(* IEC 61131-3 sources: NachHouse_TST/ROOM_API_PILOT/CODEX_BACKUP_BEFORE_SORT_FIX_20260827_0827, 1 file *)

(* ---- 08_COMMAND_ENGINE.ST ---- *)
(* Spracovanie príkazov ADD / DELETE / COPY / SET pre miestnosti. ENG *)

(* Spracuje najviac jeden príkaz, iba ak klient nastavil ApiCommandExecute. *)
FUNCTION ApiProcessRoomCommand : BOOL
VAR
    i             : USINT;     (* Index pri prechode poľom miestností. *)
    configSlot    : USINT;     (* Nájdená alebo voľná pozícia cieľovej konfigurácie. ENG *)
    stateSlot     : USINT;     (* Nájdená alebo voľná pozícia cieľového stavu. ENG *)
    sourceCfgSlot : USINT;     (* Pozícia zdrojovej konfigurácie pri kopírovaní. ENG *)
    sourceStSlot  : USINT;     (* Pozícia zdrojového stavu pri kopírovaní. ENG *)
    maxSort       : UINT;      (* Najvyššie použité predvolené poradie pri pridávaní. ENG *)
    sourceSort    : UINT;      (* Predvolené poradie zdroja pri vkladaní jeho kópie. ENG *)
    resultCode    : USINT;     (* Pracovný návratový kód API_RESULT_*. ENG *)
    resultMessage : STRING[80]; (* Pracovný slovenský text výsledku. *)
    executeChange : BOOL;      (* TRUE iba vtedy, keď sa snapshot skutočne zmenil. ENG *)
END_VAR

(* Bez spúšťacieho príznaku funkcia okamžite skončí bez vedľajších účinkov. *)
ApiProcessRoomCommand := FALSE;
IF NOT ApiCommandExecute THEN
    RETURN;
END_IF;

(* Začiatok dvojfázového handshake: príkaz je prevzatý na spracovanie. ENG *)
ApiProcessRoomCommand := TRUE;
ApiCommandBusy := TRUE;
ApiCommandFinished := FALSE;

(* Presné zopakovanie posledného ClientId + RequestId je idempotentné. ENG *)
IF (ApiCommandRoom.ClientId = ApiLastCommandClientId) AND
   (ApiCommandRoom.RequestId = ApiLastCommandRequestId) AND
   (ApiCommandRoom.RequestId <> 0) THEN

    ApiCommandResult := ApiLastStoredResult;
    ApiInfo.LastCommandResult := ApiLastStoredResult;

ELSE
    (* Predvolené hodnoty pre nový, ešte nespracovaný príkaz. *)
    resultCode := API_RESULT_OK;
    resultMessage := 'OK';
    executeChange := FALSE;

    (* Spoločná kontrola povinných identifikátorov transportu. *)
    IF (ApiCommandRoom.ClientId = '') OR (ApiCommandRoom.RequestId = 0) THEN
        resultCode := API_RESULT_INVALID_ARGUMENT;
        resultMessage := 'Neplatny ClientId alebo RequestId';
    ELSE
        (* Rozdelenie spracovania podľa verejného číselného kódu Action. ENG *)
        CASE ApiCommandRoom.Action OF

            API_ACTION_ADD_ROOM:
                (* ADD: overí cieľ, nájde voľné sloty a vytvorí konfiguráciu aj stav. ENG *)
                IF (ApiCommandRoom.RoomId = 0) OR (ApiCommandRoom.Name = '') THEN
                    resultCode := API_RESULT_INVALID_ARGUMENT;
                    resultMessage := 'Neplatne ID alebo nazov';
                ELSIF ApiFindConfigSlot(ApiCommandRoom.RoomId) <> 0 THEN
                    resultCode := API_RESULT_ALREADY_EXISTS;
                    resultMessage := 'RoomId uz existuje';
                ELSE
                    configSlot := ApiFindFreeConfigSlot();
                    stateSlot := ApiFindFreeStateSlot();
                    IF (configSlot = 0) OR (stateSlot = 0) THEN
                        resultCode := API_RESULT_NO_FREE_SLOT;
                        resultMessage := 'Nie je volny slot';
                    ELSE
                        (* Nová miestnosť sa zaradí za najvyššie existujúce SortDefault. ENG *)
                        maxSort := 0;
                        FOR i := 1 TO C_MAX_ROOMS DO
                            IF ApiConfig.Rooms[i].Used AND
                               (ApiConfig.Rooms[i].SortDefault > maxSort) THEN
                                maxSort := ApiConfig.Rooms[i].SortDefault;
                            END_IF;
                        END_FOR;

                        (* Vytvorenie cieľovej konfigurácie z údajov klienta a predvolenej ikony. *)
                        ApiClearRoomConfig(ApiConfig.Rooms[configSlot]);
                        ApiConfig.Rooms[configSlot].Used := TRUE;
                        ApiConfig.Rooms[configSlot].RoomId := ApiCommandRoom.RoomId;
                        ApiConfig.Rooms[configSlot].Name := ApiCommandRoom.Name;
                        ApiConfig.Rooms[configSlot].ProjectName := ApiCommandRoom.ProjectName;
                        ApiConfig.Rooms[configSlot].IconId := API_DEFAULT_ICON_ID;
                        ApiConfig.Rooms[configSlot].SortDefault := maxSort + 1;

                        (* Vytvorenie samostatného stavového záznamu s testovacími hodnotami. *)
                        ApiClearRoomState(ApiState.Rooms[stateSlot]);
                        ApiState.Rooms[stateSlot].RoomId := ApiCommandRoom.RoomId;
                        ApiState.Rooms[stateSlot].Temperature := API_DEFAULT_TEMPERATURE;
                        ApiState.Rooms[stateSlot].Humidity := API_DEFAULT_HUMIDITY;
                        ApiState.Rooms[stateSlot].Presence := FALSE;
                        ApiState.Rooms[stateSlot].DayPhase := API_DAY_PHASE_DAY;
                        ApiState.Rooms[stateSlot].CategoryMask := DWORD#16#00000000;
                        ApiState.Rooms[stateSlot].AlarmLevel := API_ALARM_OK;
                        ApiState.Rooms[stateSlot].Online := TRUE;

                        executeChange := TRUE;
                        resultMessage := 'Miestnost pridana';
                    END_IF;
                END_IF;

            API_ACTION_DELETE_ROOM:
                (* DELETE: konfigurácia aj stav musia existovať, potom sa oba sloty vyčistia. ENG *)
                configSlot := ApiFindConfigSlot(ApiCommandRoom.RoomId);
                stateSlot := ApiFindStateSlot(ApiCommandRoom.RoomId);
                IF (configSlot = 0) OR (stateSlot = 0) THEN
                    resultCode := API_RESULT_NOT_FOUND;
                    resultMessage := 'Miestnost nenajdena';
                ELSE
                    ApiClearRoomConfig(ApiConfig.Rooms[configSlot]);
                    ApiClearRoomState(ApiState.Rooms[stateSlot]);
                    executeChange := TRUE;
                    resultMessage := 'Miestnost zmazana';
                END_IF;

            API_ACTION_COPY_ROOM:
                (* COPY: najprv sa overí zdroj aj jedinečnosť cieľového RoomId. ENG *)
                sourceCfgSlot := ApiFindConfigSlot(ApiCommandRoom.SourceRoomId);
                sourceStSlot := ApiFindStateSlot(ApiCommandRoom.SourceRoomId);
                IF (ApiCommandRoom.RoomId = 0) OR
                   (ApiCommandRoom.RoomId = ApiCommandRoom.SourceRoomId) THEN
                    resultCode := API_RESULT_INVALID_ARGUMENT;
                    resultMessage := 'Neplatne cielove RoomId';
                ELSIF (sourceCfgSlot = 0) OR (sourceStSlot = 0) THEN
                    resultCode := API_RESULT_NOT_FOUND;
                    resultMessage := 'Zdrojova miestnost nenajdena';
                ELSIF ApiFindConfigSlot(ApiCommandRoom.RoomId) <> 0 THEN
                    resultCode := API_RESULT_ALREADY_EXISTS;
                    resultMessage := 'Cielove RoomId uz existuje';
                ELSE
                    configSlot := ApiFindFreeConfigSlot();
                    stateSlot := ApiFindFreeStateSlot();
                    IF (configSlot = 0) OR (stateSlot = 0) THEN
                        resultCode := API_RESULT_NO_FREE_SLOT;
                        resultMessage := 'Nie je volny slot';
                    ELSE
                        (* Pre kópiu sa uvoľní poradie hneď za zdrojovou miestnosťou. *)
                        sourceSort := ApiConfig.Rooms[sourceCfgSlot].SortDefault;
                        FOR i := 1 TO C_MAX_ROOMS DO
                            IF ApiConfig.Rooms[i].Used AND
                               (ApiConfig.Rooms[i].SortDefault > sourceSort) THEN
                                ApiConfig.Rooms[i].SortDefault :=
                                    ApiConfig.Rooms[i].SortDefault + 1;
                            END_IF;
                        END_FOR;

                        (* Konfigurácia sa kopíruje celá; klient môže voliteľne prepísať názvy. *)
                        ApiConfig.Rooms[configSlot] := ApiConfig.Rooms[sourceCfgSlot];
                        ApiConfig.Rooms[configSlot].RoomId := ApiCommandRoom.RoomId;
                        ApiConfig.Rooms[configSlot].SortDefault := sourceSort + 1;
                        IF ApiCommandRoom.Name <> '' THEN
                            ApiConfig.Rooms[configSlot].Name := ApiCommandRoom.Name;
                        END_IF;
                        IF ApiCommandRoom.ProjectName <> '' THEN
                            ApiConfig.Rooms[configSlot].ProjectName := ApiCommandRoom.ProjectName;
                        END_IF;

                        (* Pilot kopíruje aj ručne nastavený stav, ale priradí nové RoomId. ENG *)
                        ApiState.Rooms[stateSlot] := ApiState.Rooms[sourceStSlot];
                        ApiState.Rooms[stateSlot].RoomId := ApiCommandRoom.RoomId;

                        executeChange := TRUE;
                        resultMessage := 'Miestnost skopirovana';
                    END_IF;
                END_IF;

            API_ACTION_SET_ROOM_DATA:
                (* SET: v pilote mení iba hlavný a doplnkový názov miestnosti. ENG *)
                configSlot := ApiFindConfigSlot(ApiCommandRoom.RoomId);
                IF configSlot = 0 THEN
                    resultCode := API_RESULT_NOT_FOUND;
                    resultMessage := 'Miestnost nenajdena';
                ELSIF ApiCommandRoom.Name = '' THEN
                    resultCode := API_RESULT_INVALID_ARGUMENT;
                    resultMessage := 'Nazov nesmie byt prazdny';
                ELSE
                    ApiConfig.Rooms[configSlot].Name := ApiCommandRoom.Name;
                    ApiConfig.Rooms[configSlot].ProjectName := ApiCommandRoom.ProjectName;
                    executeChange := TRUE;
                    resultMessage := 'Udaje miestnosti nastavene';
                END_IF;

            ELSE
                (* Neznámy číselný kód Action sa odmietne bez zmeny dát. ENG *)
                resultCode := API_RESULT_UNSUPPORTED_ACTION;
                resultMessage := 'Nepodporovana akcia';
        END_CASE;
    END_IF;

    (* Úspešná dátová zmena vytvorí nové revízie a príslušné diff rámce. ENG *)
    IF executeChange AND (resultCode = API_RESULT_OK) THEN
        ApiCaptureConfigChanges();
        ApiCaptureStateChanges();
    END_IF;

    (* Výsledok nesie identitu požiadavky aj revízie platné po jej spracovaní. *)
    ApiCommandResult.ClientId := ApiCommandRoom.ClientId;
    ApiCommandResult.RequestId := ApiCommandRoom.RequestId;
    ApiCommandResult.Result := resultCode;
    ApiCommandResult.Message := resultMessage;
    ApiCommandResult.ConfigRevision := ApiInfo.ConfigRevision;
    ApiCommandResult.StateRevision := ApiInfo.StateRevision;

    (* Uloženie výsledku pre ApiInfo a idempotentné opakovanie poslednej požiadavky. *)
    ApiInfo.LastCommandResult := ApiCommandResult;
    ApiLastCommandClientId := ApiCommandRoom.ClientId;
    ApiLastCommandRequestId := ApiCommandRoom.RequestId;
    ApiLastStoredResult := ApiCommandResult;
END_IF;

(* Ukončenie handshake: PLC zruší Execute, uvoľní Busy a nastaví Finished. ENG *)
ApiCommandExecute := FALSE;
ApiCommandBusy := FALSE;
ApiCommandFinished := TRUE;
END_FUNCTION
